TYPE stMessageFormat :
STRUCT
	sDateTime							: STRING[25];
	sErrID								: STRING[11];
	sLevel								: STRING[10];
	sModuleDescription					: STRING[80];
	sErrorMessage						: STRING[200];	
END_STRUCT
END_TYPE

(* stored: Version 1.1.0.1, ProductVersion 3.1.4024.13
   DUT stMessageFormat: Id {ad740de9-e962-443d-9685-e65bb54a1a7a} *)
